(* PLC project counter, tcpethernet counter 1 *)
(* stored: creationDateTime 2026-10-28T09:00:00, modificationDateTime 2026-10-28T09:00:00 *)

PROGRAM counter
  VAR
    Pulse AT %IX0.2 : BOOL;
    Reset AT %IX0.3 : BOOL;
  END_VAR
  VAR CONSTANT
    Limit : INT := 3;
  END_VAR
  VAR
    count : INT;
    Done : BOOL;
    AtMostOne : BOOL;
    ctr : CTU;
  END_VAR

(* FBD diagram, written out as Structured Text *)
ctr(CU := Pulse, R := Reset, PV := Limit);
Done := ctr.Q;
count := ctr.CV;
AtMostOne := NOT (ctr.CV > 1);
(* AtMostOne is NOT (count > 1) *)
END_PROGRAM
